// TIA Portal project "PRODUCTION_CIMENT" (V16)

(* hardware
DEVICE "Station S7-1200_1"  S7-1200 Station
   slot 0: "Châssis_0"  S7-1200 Rack  Rack  V1.0
   slot 1: "PLC_1"  CPU 1214C AC/DC/Rly  6ES7 214-1BG40-0XB0  V4.4
*)

// ===== PLC "PLC_1"  CPU 1214C AC/DC/Rly =====

VAR_GLOBAL   // PLC tag table "Table de variables standard"
   "Tag_1" AT %M0.1 : Bool;
   "X0" AT %M0.2 : Bool;
   "X1" AT %M0.3 : Bool;
   "STOP" AT %I0.0 : Bool;
   "START" AT %I0.1 : Bool;
   "X20" AT %M0.4 : Bool;
   "X21" AT %M1.0 : Bool;
   "X22" AT %M1.1 : Bool;
   "X23" AT %M1.2 : Bool;
   "X24" AT %M1.3 : Bool;
   "BP_Reset" AT %I0.2 : Bool;
   "BP_Marche" AT %I0.3 : Bool;
   "Cap_Niveau_Tremie" AT %I0.4 : Bool;
   "Cap_Pression" AT %I0.5 : Bool;
   "Detect_Blocage" AT %I0.6 : Bool;
   "Cap_Charge_Moteur" AT %I0.7 : Bool;
   "Memo_T1" AT %MD1 : Time;
   "Cap_Vitesse" AT %I1.0 : Bool;
   "KM1" AT %Q0.1 : Bool;
   "Concasseur" AT %Q0.2 : Bool;
   "X30" AT %M1.4 : Bool;
   "X31" AT %M1.5 : Bool;
   "X32" AT %M1.6 : Bool;
   "X33" AT %M1.7 : Bool;
   "X34" AT %M2.0 : Bool;
   "Bp_Reset2" AT %I1.1 : Bool;
   "Cap_Portes" AT %I1.3 : Bool;
   "Cap_Vibration" AT %I1.4 : Bool;
   "Cap_Temperature" AT %I1.5 : Bool;
   "Cap_Vitesse2" AT %I1.6 : Bool;
   "Cap_Charge2" AT %I1.7 : Bool;
   "Cap_Pression2" AT %I2.0 : Bool;
   "Detect_Corps_Etrangers" AT %I2.1 : Bool;
   "Cap_Debit" AT %I2.2 : Bool;
   "BP_Marche_Concasseur_Sec" AT %I2.3 : Bool;
   "Cap_Niveau2" AT %I2.4 : Bool;
   "SAU1" AT %I2.5 : Bool;
   "KM2" AT %Q0.3 : Bool;
   "Concasseur2" AT %Q0.4 : Bool;
   "X40" AT %M2.1 : Bool;
   "X41" AT %M2.2 : Bool;
   "X42" AT %M2.3 : Bool;
   "X43" AT %M2.4 : Bool;
   "X44" AT %M2.5 : Bool;
   "X45" AT %M2.6 : Bool;
   "X46" AT %M2.7 : Bool;
   "X47" AT %M3.0 : Bool;
   "BP_Reset3" AT %I2.6 : Bool;
   "BP_Marche_Broyeur" AT %I2.7 : Bool;
   "Cap_Niveau_Mat" AT %I3.0 : Bool;
   "Cap_Temperature_Paliers" AT %I3.1 : Bool;
   "Cap_Vitesse_Broyeur" AT %I3.2 : Bool;
   "BP_Stop_Broyeur" AT %I3.3 : Bool;
   "MemoT2" AT %MD3 : Time;
END_VAR

// folder: System blocks/Program resources

DATA_BLOCK "T1"   // DB1
{ S7_Optimized_Access := 'TRUE' }
AUTHOR : Simatic
FAMILY : IEC
NAME : IEC_TMR
VERSION : 1.0
// stored: InstanceOfName IEC_TIMER
"IEC_TIMER"
BEGIN
END_DATA_BLOCK

DATA_BLOCK "T2"   // DB2
{ S7_Optimized_Access := 'TRUE' }
AUTHOR : Simatic
FAMILY : IEC
NAME : IEC_TMR
VERSION : 1.0
// stored: InstanceOfName IEC_TIMER
"IEC_TIMER"
BEGIN
END_DATA_BLOCK

DATA_BLOCK "T3"   // DB3
{ S7_Optimized_Access := 'TRUE' }
AUTHOR : Simatic
FAMILY : IEC
NAME : IEC_TMR
VERSION : 1.0
// stored: InstanceOfName IEC_TIMER
"IEC_TIMER"
BEGIN
END_DATA_BLOCK

// folder: (top level)

FUNCTION_BLOCK "GC"   // FB1, LAD
{ S7_Optimized_Access := 'TRUE' }
VERSION : 0.1
BEGIN

REGION Network 1
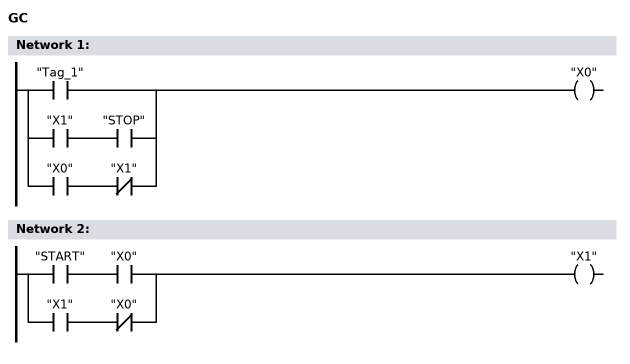
   RUNG wire#powerrail
      Contact( "Tag_1" )
      wire#w1
      Coil( "X0" )
   END_RUNG
   RUNG wire#powerrail
      Contact( "X1" )
      Contact( "STOP" )
   END_RUNG wire#w1
   RUNG wire#powerrail
      Contact( "X0" )
      I_Contact( "X1" )
   END_RUNG wire#w1
   // the same network as SCL:
   "X0" := "Tag_1" OR ("X1" AND "STOP") OR ("X0" AND NOT "X1");
END_REGION

REGION Network 2
   RUNG wire#powerrail
      Contact( "START" )
      Contact( "X0" )
      wire#w1
      Coil( "X1" )
   END_RUNG
   RUNG wire#powerrail
      Contact( "X1" )
      I_Contact( "X0" )
   END_RUNG wire#w1
   // the same network as SCL:
   "X1" := ("START" AND "X0") OR ("X1" AND NOT "X0");
END_REGION
END_FUNCTION_BLOCK

FUNCTION_BLOCK "GFN"   // FB2, LAD
{ S7_Optimized_Access := 'TRUE' }
VERSION : 0.1
BEGIN
END_FUNCTION_BLOCK

FUNCTION_BLOCK "GT1"   // FB3, LAD
{ S7_Optimized_Access := 'TRUE' }
VERSION : 0.1
BEGIN

REGION Network 1
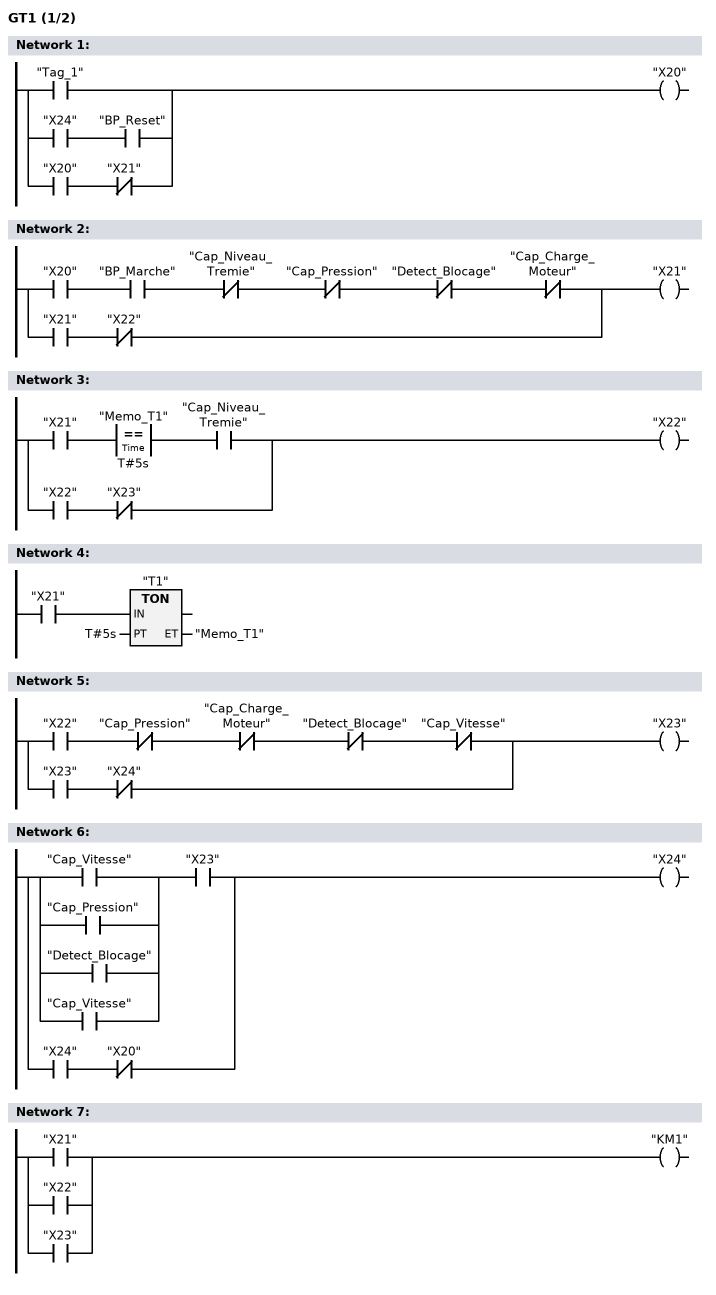
   RUNG wire#powerrail
      Contact( "Tag_1" )
      wire#w1
      Coil( "X20" )
   END_RUNG
   RUNG wire#powerrail
      Contact( "X24" )
      Contact( "BP_Reset" )
   END_RUNG wire#w1
   RUNG wire#powerrail
      Contact( "X20" )
      I_Contact( "X21" )
   END_RUNG wire#w1
   // the same network as SCL:
   "X20" := "Tag_1" OR ("X24" AND "BP_Reset") OR ("X20" AND NOT "X21");
END_REGION

REGION Network 2
   RUNG wire#powerrail
      Contact( "X20" )
      Contact( "BP_Marche" )
      I_Contact( "Cap_Niveau_Tremie" )
      I_Contact( "Cap_Pression" )
      I_Contact( "Detect_Blocage" )
      I_Contact( "Cap_Charge_Moteur" )
      wire#w1
      Coil( "X21" )
   END_RUNG
   RUNG wire#powerrail
      Contact( "X21" )
      I_Contact( "X22" )
   END_RUNG wire#w1
   // the same network as SCL:
   "X21" := ("X20" AND "BP_Marche" AND NOT "Cap_Niveau_Tremie" AND NOT "Cap_Pression" AND NOT "Detect_Blocage" AND NOT "Cap_Charge_Moteur") OR ("X21" AND NOT "X22");
END_REGION

REGION Network 3
   RUNG wire#powerrail
      Contact( "X21" )
      { S7_Templates := "SrcType := Time" } EQ_Contact(in1 := "Memo_T1", in2 := T#5s)
      Contact( "Cap_Niveau_Tremie" )
      wire#w1
      Coil( "X22" )
   END_RUNG
   RUNG wire#powerrail
      Contact( "X22" )
      I_Contact( "X23" )
   END_RUNG wire#w1
   // the same network as SCL:
   "X22" := ("X21" AND ("Memo_T1" = T#5s) AND "Cap_Niveau_Tremie") OR ("X22" AND NOT "X23");
END_REGION

REGION Network 4
   "T1".TON(IN := "X21", PT := T#5s, ET => "Memo_T1");
END_REGION

REGION Network 5
   RUNG wire#powerrail
      Contact( "X22" )
      I_Contact( "Cap_Pression" )
      I_Contact( "Cap_Charge_Moteur" )
      I_Contact( "Detect_Blocage" )
      I_Contact( "Cap_Vitesse" )
      wire#w1
      Coil( "X23" )
   END_RUNG
   RUNG wire#powerrail
      Contact( "X23" )
      I_Contact( "X24" )
   END_RUNG wire#w1
   // the same network as SCL:
   "X23" := ("X22" AND NOT "Cap_Pression" AND NOT "Cap_Charge_Moteur" AND NOT "Detect_Blocage" AND NOT "Cap_Vitesse") OR ("X23" AND NOT "X24");
END_REGION

REGION Network 6
   RUNG wire#powerrail
      Contact( "Cap_Vitesse" )
      wire#w1
      Contact( "X23" )
      wire#w2
      Coil( "X24" )
   END_RUNG
   RUNG wire#powerrail
      Contact( "Cap_Pression" )
   END_RUNG wire#w1
   RUNG wire#powerrail
      Contact( "Detect_Blocage" )
   END_RUNG wire#w1
   RUNG wire#powerrail
      Contact( "Cap_Vitesse" )
   END_RUNG wire#w1
   RUNG wire#powerrail
      Contact( "X24" )
      I_Contact( "X20" )
   END_RUNG wire#w2
   // the same network as SCL:
   "X24" := (("Cap_Vitesse" OR "Cap_Pression" OR "Detect_Blocage" OR "Cap_Vitesse") AND "X23") OR ("X24" AND NOT "X20");
END_REGION

REGION Network 7
   RUNG wire#powerrail
      Contact( "X21" )
      wire#w1
      Coil( "KM1" )
   END_RUNG
   RUNG wire#powerrail
      Contact( "X22" )
   END_RUNG wire#w1
   RUNG wire#powerrail
      Contact( "X23" )
   END_RUNG wire#w1
   // the same network as SCL:
   "KM1" := "X21" OR "X22" OR "X23";
END_REGION

REGION Network 8
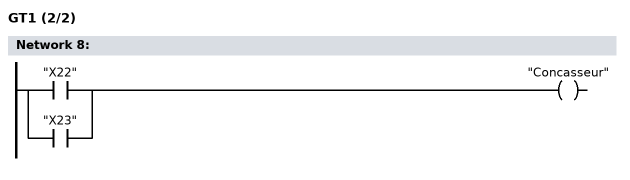
   RUNG wire#powerrail
      Contact( "X22" )
      wire#w1
      Coil( "Concasseur" )
   END_RUNG
   RUNG wire#powerrail
      Contact( "X23" )
   END_RUNG wire#w1
   // the same network as SCL:
   "Concasseur" := "X22" OR "X23";
END_REGION
END_FUNCTION_BLOCK

FUNCTION_BLOCK "GT2"   // FB4, LAD
{ S7_Optimized_Access := 'TRUE' }
VERSION : 0.1
// GRAFCET DE TACHE 2, CONCASSEUR SECONDAIRE
BEGIN

REGION Network 1: ETAPE 30
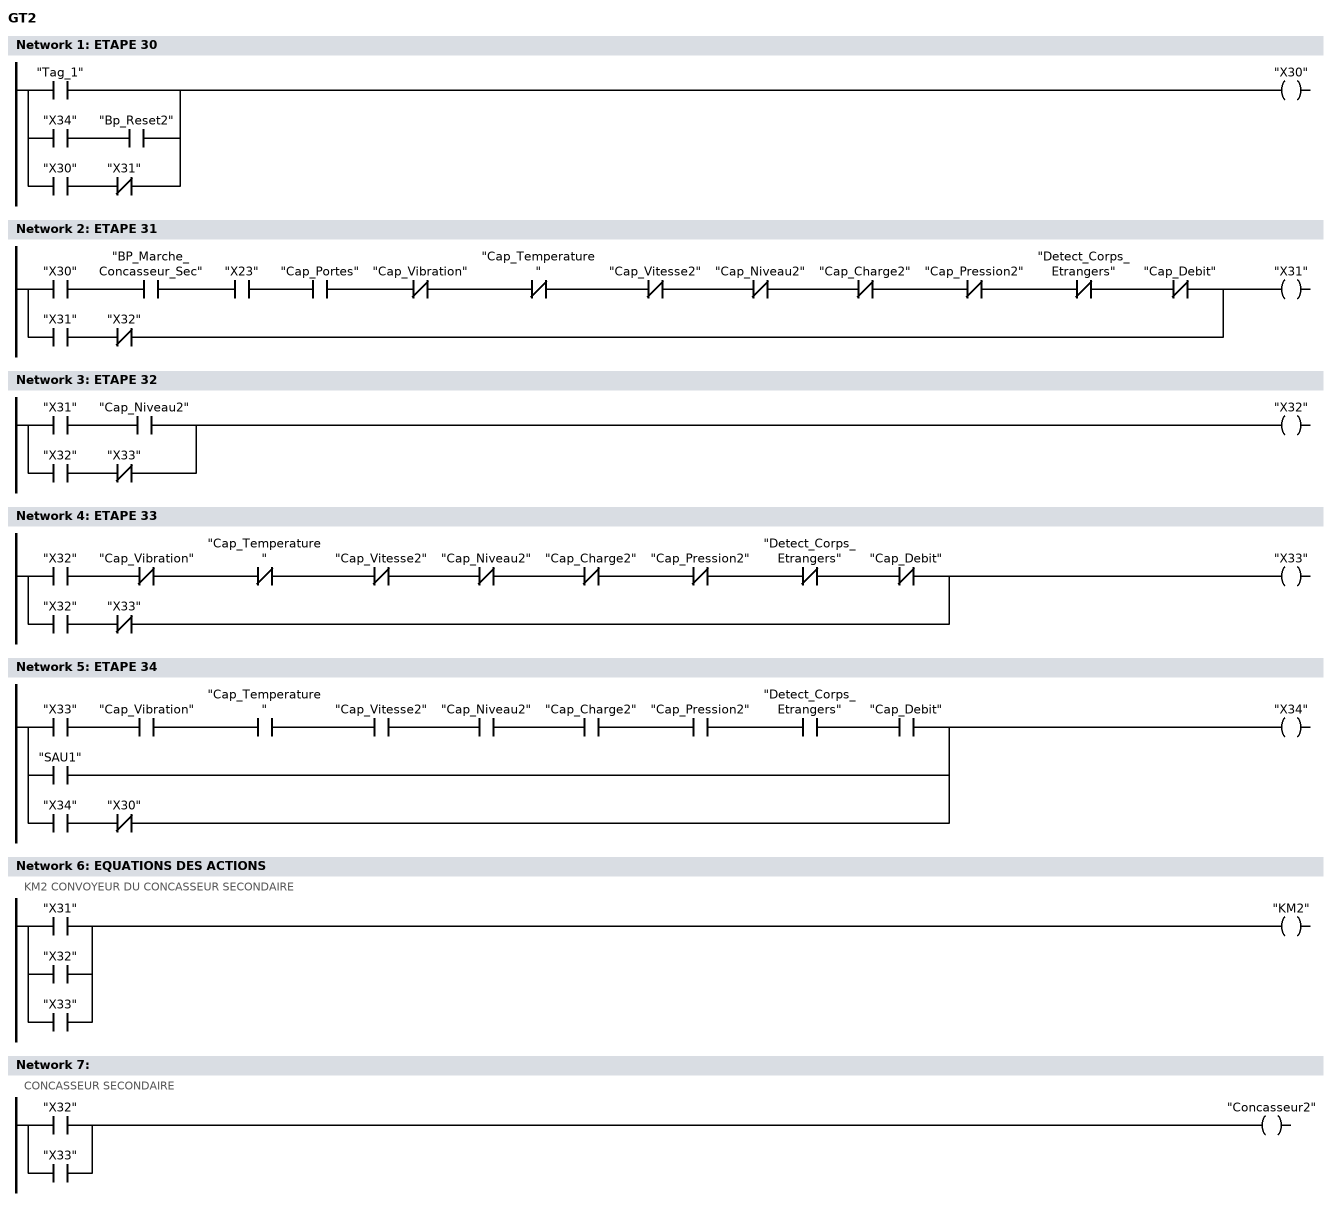
   RUNG wire#powerrail
      Contact( "Tag_1" )
      wire#w1
      Coil( "X30" )
   END_RUNG
   RUNG wire#powerrail
      Contact( "X34" )
      Contact( "Bp_Reset2" )
   END_RUNG wire#w1
   RUNG wire#powerrail
      Contact( "X30" )
      I_Contact( "X31" )
   END_RUNG wire#w1
   // the same network as SCL:
   "X30" := "Tag_1" OR ("X34" AND "Bp_Reset2") OR ("X30" AND NOT "X31");
END_REGION

REGION Network 2: ETAPE 31
   RUNG wire#powerrail
      Contact( "X30" )
      Contact( "BP_Marche_Concasseur_Sec" )
      Contact( "X23" )
      Contact( "Cap_Portes" )
      I_Contact( "Cap_Vibration" )
      I_Contact( "Cap_Temperature" )
      I_Contact( "Cap_Vitesse2" )
      I_Contact( "Cap_Niveau2" )
      I_Contact( "Cap_Charge2" )
      I_Contact( "Cap_Pression2" )
      I_Contact( "Detect_Corps_Etrangers" )
      I_Contact( "Cap_Debit" )
      wire#w1
      Coil( "X31" )
   END_RUNG
   RUNG wire#powerrail
      Contact( "X31" )
      I_Contact( "X32" )
   END_RUNG wire#w1
   // the same network as SCL:
   "X31" := ("X30" AND "BP_Marche_Concasseur_Sec" AND "X23" AND "Cap_Portes" AND NOT "Cap_Vibration" AND NOT "Cap_Temperature" AND NOT "Cap_Vitesse2" AND NOT "Cap_Niveau2" AND NOT "Cap_Charge2" AND NOT "Cap_Pression2" AND NOT "Detect_Corps_Etrangers" AND NOT "Cap_Debit") OR ("X31" AND NOT "X32");
END_REGION

REGION Network 3: ETAPE 32
   RUNG wire#powerrail
      Contact( "X31" )
      Contact( "Cap_Niveau2" )
      wire#w1
      Coil( "X32" )
   END_RUNG
   RUNG wire#powerrail
      Contact( "X32" )
      I_Contact( "X33" )
   END_RUNG wire#w1
   // the same network as SCL:
   "X32" := ("X31" AND "Cap_Niveau2") OR ("X32" AND NOT "X33");
END_REGION

REGION Network 4: ETAPE 33
   RUNG wire#powerrail
      Contact( "X32" )
      I_Contact( "Cap_Vibration" )
      I_Contact( "Cap_Temperature" )
      I_Contact( "Cap_Vitesse2" )
      I_Contact( "Cap_Niveau2" )
      I_Contact( "Cap_Charge2" )
      I_Contact( "Cap_Pression2" )
      I_Contact( "Detect_Corps_Etrangers" )
      I_Contact( "Cap_Debit" )
      wire#w1
      Coil( "X33" )
   END_RUNG
   RUNG wire#powerrail
      Contact( "X32" )
      I_Contact( "X33" )
   END_RUNG wire#w1
   // the same network as SCL:
   "X33" := ("X32" AND NOT "Cap_Vibration" AND NOT "Cap_Temperature" AND NOT "Cap_Vitesse2" AND NOT "Cap_Niveau2" AND NOT "Cap_Charge2" AND NOT "Cap_Pression2" AND NOT "Detect_Corps_Etrangers" AND NOT "Cap_Debit") OR ("X32" AND NOT "X33");
END_REGION

REGION Network 5: ETAPE 34
   RUNG wire#powerrail
      Contact( "X33" )
      Contact( "Cap_Vibration" )
      Contact( "Cap_Temperature" )
      Contact( "Cap_Vitesse2" )
      Contact( "Cap_Niveau2" )
      Contact( "Cap_Charge2" )
      Contact( "Cap_Pression2" )
      Contact( "Detect_Corps_Etrangers" )
      Contact( "Cap_Debit" )
      wire#w1
      Coil( "X34" )
   END_RUNG
   RUNG wire#powerrail
      Contact( "SAU1" )
   END_RUNG wire#w1
   RUNG wire#powerrail
      Contact( "X34" )
      I_Contact( "X30" )
   END_RUNG wire#w1
   // the same network as SCL:
   "X34" := ("X33" AND "Cap_Vibration" AND "Cap_Temperature" AND "Cap_Vitesse2" AND "Cap_Niveau2" AND "Cap_Charge2" AND "Cap_Pression2" AND "Detect_Corps_Etrangers" AND "Cap_Debit") OR "SAU1" OR ("X34" AND NOT "X30");
END_REGION

REGION Network 6: EQUATIONS DES ACTIONS
   // KM2 CONVOYEUR DU CONCASSEUR SECONDAIRE
   RUNG wire#powerrail
      Contact( "X31" )
      wire#w1
      Coil( "KM2" )
   END_RUNG
   RUNG wire#powerrail
      Contact( "X32" )
   END_RUNG wire#w1
   RUNG wire#powerrail
      Contact( "X33" )
   END_RUNG wire#w1
   // the same network as SCL:
   "KM2" := "X31" OR "X32" OR "X33";
END_REGION

REGION Network 7
   // CONCASSEUR SECONDAIRE
   RUNG wire#powerrail
      Contact( "X32" )
      wire#w1
      Coil( "Concasseur2" )
   END_RUNG
   RUNG wire#powerrail
      Contact( "X33" )
   END_RUNG wire#w1
   // the same network as SCL:
   "Concasseur2" := "X32" OR "X33";
END_REGION
END_FUNCTION_BLOCK

FUNCTION_BLOCK "GT3"   // FB5, LAD
{ S7_Optimized_Access := 'TRUE' }
VERSION : 0.1
// GRAFCET  DE TACHE 3 BROYEUR :
BEGIN

REGION Network 1: EQUATIONS DES ETAPES
   // ETAPE X40
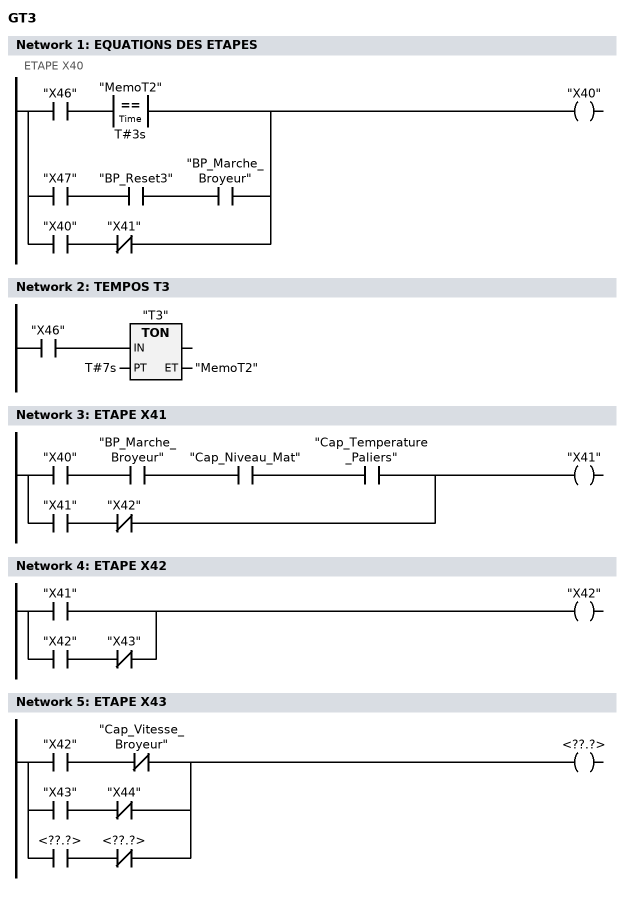
   RUNG wire#powerrail
      Contact( "X46" )
      { S7_Templates := "SrcType := Time" } EQ_Contact(in1 := "MemoT2", in2 := T#3s)
      wire#w1
      Coil( "X40" )
   END_RUNG
   RUNG wire#powerrail
      Contact( "X47" )
      Contact( "BP_Reset3" )
      Contact( "BP_Marche_Broyeur" )
   END_RUNG wire#w1
   RUNG wire#powerrail
      Contact( "X40" )
      I_Contact( "X41" )
   END_RUNG wire#w1
   // the same network as SCL:
   "X40" := ("X46" AND ("MemoT2" = T#3s)) OR ("X47" AND "BP_Reset3" AND "BP_Marche_Broyeur") OR ("X40" AND NOT "X41");
END_REGION

REGION Network 2: TEMPOS T3
   "T3".TON(IN := "X46", PT := T#7s, ET => "MemoT2");
END_REGION

REGION Network 3: ETAPE X41
   RUNG wire#powerrail
      Contact( "X40" )
      Contact( "BP_Marche_Broyeur" )
      Contact( "Cap_Niveau_Mat" )
      Contact( "Cap_Temperature_Paliers" )
      wire#w1
      Coil( "X41" )
   END_RUNG
   RUNG wire#powerrail
      Contact( "X41" )
      I_Contact( "X42" )
   END_RUNG wire#w1
   // the same network as SCL:
   "X41" := ("X40" AND "BP_Marche_Broyeur" AND "Cap_Niveau_Mat" AND "Cap_Temperature_Paliers") OR ("X41" AND NOT "X42");
END_REGION

REGION Network 4: ETAPE X42
   RUNG wire#powerrail
      Contact( "X41" )
      wire#w1
      Coil( "X42" )
   END_RUNG
   RUNG wire#powerrail
      Contact( "X42" )
      I_Contact( "X43" )
   END_RUNG wire#w1
   // the same network as SCL:
   "X42" := "X41" OR ("X42" AND NOT "X43");
END_REGION

REGION Network 5: ETAPE X43
   RUNG wire#powerrail
      Contact( "X42" )
      I_Contact( "Cap_Vitesse_Broyeur" )
      wire#w1
      Coil(  )
   END_RUNG
   RUNG wire#powerrail
      Contact( "X43" )
      I_Contact( "X44" )
   END_RUNG wire#w1
   RUNG wire#powerrail
      Contact(  )
      I_Contact(  )
   END_RUNG wire#w1
   // the same network as SCL:
   // no checked SCL form for this network; see the picture
END_REGION
END_FUNCTION_BLOCK

ORGANIZATION_BLOCK "Main"   // OB1, LAD, ProgramCycle
TITLE = "Main Program Sweep (Cycle)"
{ S7_Optimized_Access := 'TRUE' }
VERSION : 0.1
   VAR_INPUT
      Initial_Call : Bool;   // Initial call of this OB
      Remanence : Bool;   // =True, if remanent data are available
   END_VAR
BEGIN
END_ORGANIZATION_BLOCK